PROGRAM MAIN

VAR CONSTANT 
    deviceCount : WORD := 3;
END_VAR

VAR
	// Outputs
	{attribute 'TcLinkTo' := '[1].mDirection := TIID^Device_1^Box 1 (LAN9255_EtherCAT_Slave)^Outputs process data mapping^Direction;
								[1].mSpeed := TIID^Device_1^Box 1 (LAN9255_EtherCAT_Slave)^Outputs process data mapping^Speed;
								[1].mTime := TIID^Device_1^Box 1 (LAN9255_EtherCAT_Slave)^Outputs process data mapping^Time;
								[1].mMode := TIID^Device_1^Box 1 (LAN9255_EtherCAT_Slave)^Outputs process data mapping^Mode;
								
								[2].mDirection := TIID^Device_1^Box 2 (LAN9255_EtherCAT_Slave)^Outputs process data mapping^Direction;
								[2].mSpeed := TIID^Device_1^Box 2 (LAN9255_EtherCAT_Slave)^Outputs process data mapping^Speed;
								[2].mTime := TIID^Device_1^Box 2 (LAN9255_EtherCAT_Slave)^Outputs process data mapping^Time;
								[2].mMode := TIID^Device_1^Box 2 (LAN9255_EtherCAT_Slave)^Outputs process data mapping^Mode;
								
								[3].mDirection := TIID^Device_1^Box 3 (LAN9255_EtherCAT_Slave)^Outputs process data mapping^Direction;
								[3].mSpeed := TIID^Device_1^Box 3 (LAN9255_EtherCAT_Slave)^Outputs process data mapping^Speed;
								[3].mTime := TIID^Device_1^Box 3 (LAN9255_EtherCAT_Slave)^Outputs process data mapping^Time;
								[3].mMode := TIID^Device_1^Box 3 (LAN9255_EtherCAT_Slave)^Outputs process data mapping^Mode'}
	device : ARRAY [1..deviceCount] OF EthercatDevice ;

	// Inputs
	{attribute 'TcLinkTo' := '[1]:= TIID^Device_1^Box 1 (LAN9255_EtherCAT_Slave)^Inputs process data mapping^Position;
								[2]	:= TIID^Device_1^Box 2 (LAN9255_EtherCAT_Slave)^Inputs process data mapping^Position;
								[3]	:= TIID^Device_1^Box 3 (LAN9255_EtherCAT_Slave)^Inputs process data mapping^Position'}
	mPosition AT %I*: ARRAY [1..deviceCount] OF DWORD ;
	
	{attribute 'TcLinkTo' := '[1]:= TIID^Device_1^Box 1 (LAN9255_EtherCAT_Slave)^Inputs process data mapping^Temperature;
								[2]	:= TIID^Device_1^Box 2 (LAN9255_EtherCAT_Slave)^Inputs process data mapping^Temperature;
								[3]	:= TIID^Device_1^Box 3 (LAN9255_EtherCAT_Slave)^Inputs process data mapping^Temperature'}
	mTemperature AT %I* : ARRAY [1..deviceCount] OF DWORD ;

	{attribute 'TcLinkTo' := '[1]:= TIID^Device_1^Box 1 (LAN9255_EtherCAT_Slave)^Inputs process data mapping^Diag1;
								[2]	:= TIID^Device_1^Box 2 (LAN9255_EtherCAT_Slave)^Inputs process data mapping^Diag1;
								[3]	:= TIID^Device_1^Box 3 (LAN9255_EtherCAT_Slave)^Inputs process data mapping^Diag1'}
	mDiag1 AT %I*: ARRAY [1..deviceCount] OF DWORD ;
	
	{attribute 'TcLinkTo' := '[1]:= TIID^Device_1^Box 1 (LAN9255_EtherCAT_Slave)^Inputs process data mapping^Diag2;
								[2]	:= TIID^Device_1^Box 2 (LAN9255_EtherCAT_Slave)^Inputs process data mapping^Diag2;
								[3]	:= TIID^Device_1^Box 3 (LAN9255_EtherCAT_Slave)^Inputs process data mapping^Diag2'}
	mDiag2 AT %I* : ARRAY [1..deviceCount] OF DWORD ;

	{attribute 'TcLinkTo' := '[1]:= TIID^Device_1^Box 1 (LAN9255_EtherCAT_Slave)^Inputs process data mapping^Diag3;
								[2]	:= TIID^Device_1^Box 2 (LAN9255_EtherCAT_Slave)^Inputs process data mapping^Diag3;
								[3]	:= TIID^Device_1^Box 3 (LAN9255_EtherCAT_Slave)^Inputs process data mapping^Diag3'}
	mDiag3 AT %I*: ARRAY [1..deviceCount] OF DWORD ;

END_VAR

END_PROGRAM

(* stored: Version 1.1.0.1, ProductVersion 3.1.4024.11
   POU MAIN: Id {6280d263-c35b-4c3c-89d3-c097ab12dca9}, SpecialFunc None *)
